(* IEC 61131-3 sources: model-first-plc-agent-ai/results/T3-W-19, 2 files *)

(* ---- a1_code.st ---- *)
FUNCTION_BLOCK TankRuntime
VAR_INPUT
    start : BOOL;
    stop : BOOL;
    LSH : BOOL;
    LSHH : BOOL;
    TON_Duration : TIME;
    TOF_Duration : TIME;
END_VAR
VAR_OUTPUT
    fill_valve : BOOL;
    discharge_valve : BOOL;
END_VAR
VAR
    active_state : INT := 0;
    next_state : INT := 0;
    filling_active : BOOL := FALSE;
    ton_q : BOOL := FALSE;
    tof_q : BOOL := FALSE;
    fill_timer : TON;
    pause_timer : TOF;
END_VAR

(* Evaluate timers using the current GRAFCET situation. *)
filling_active := (active_state = 1);

fill_timer(IN := filling_active, PT := TON_Duration);
pause_timer(IN := filling_active, PT := TOF_Duration);

ton_q := fill_timer.Q;
tof_q := pause_timer.Q;

(* Evaluate transitions from one snapshot of the active situation. *)
next_state := active_state;

CASE active_state OF
    0:
        IF start AND NOT stop AND NOT LSH AND NOT LSHH THEN
            next_state := 1;
        END_IF;

    1:
        IF stop OR LSH OR LSHH THEN
            next_state := 0;
        ELSIF ton_q AND NOT stop AND NOT LSH AND NOT LSHH THEN
            next_state := 2;
        END_IF;

    2:
        IF stop OR LSH OR LSHH THEN
            next_state := 0;
        ELSIF NOT tof_q AND NOT stop AND NOT LSH AND NOT LSHH THEN
            next_state := 1;
        END_IF;

ELSE
    next_state := 0;
END_CASE;

(* Apply the new situation to the timers immediately.
   This resets TON on leaving filling, starts the TOF off-delay
   on that same departure, and asserts TOF on entering filling.
   No further transition is evaluated during this scan. *)
IF next_state <> active_state THEN
    active_state := next_state;
    filling_active := (active_state = 1);

    fill_timer(IN := filling_active, PT := TON_Duration);
    pause_timer(IN := filling_active, PT := TOF_Duration);

    ton_q := fill_timer.Q;
    tof_q := pause_timer.Q;
END_IF;

fill_valve := (active_state = 1);
discharge_valve := FALSE;

END_FUNCTION_BLOCK

PROGRAM Main
VAR
    StartCommand AT %IX100.0 : BOOL;
    StopCommand AT %IX100.1 : BOOL;
    LSH AT %IX100.2 : BOOL;
    LSHH AT %IX100.3 : BOOL;
    FillValve AT %QX100.0 : BOOL;
    DischargeValve AT %QX100.1 : BOOL;
END_VAR
VAR
    (* Configurable commissioning defaults; adjust for the plant. *)
    TON_Duration : TIME := T#5s;
    TOF_Duration : TIME := T#5s;

    start_edge : R_TRIG;
    start : BOOL := FALSE;
    initialized : BOOL := FALSE;
    controller : TankRuntime;
END_VAR

start_edge(CLK := StartCommand);

(* Seed the edge detector without treating a held startup button
   as a new press. *)
IF NOT initialized THEN
    start := FALSE;
    initialized := TRUE;
ELSE
    start := start_edge.Q;
END_IF;

controller(
    start := start,
    stop := StopCommand,
    LSH := LSH,
    LSHH := LSHH,
    TON_Duration := TON_Duration,
    TOF_Duration := TOF_Duration
);

FillValve := controller.fill_valve;
DischargeValve := controller.discharge_valve;

END_PROGRAM

(* ---- a2_code.st ---- *)
FUNCTION_BLOCK FB_TankFilling
VAR_INPUT
    StartCommand : BOOL;
    StopCommand : BOOL;
    LSH : BOOL;
    LSHH : BOOL;
    TON_Duration : TIME;
    TOF_Duration : TIME;
END_VAR
VAR_OUTPUT
    fill_valve : BOOL;
    discharge_valve : BOOL;
END_VAR
VAR
    SequenceState : INT := 0;
    StartEdge : R_TRIG;
    FillingTON : TON;
    FillingTOF : TOF;
    start : BOOL;
    stop : BOOL;
    ton_q : BOOL;
    tof_q : BOOL;
    FillingActive : BOOL;
END_VAR

StartEdge(CLK := StartCommand);
start := StartEdge.Q;
stop := StopCommand;

(* Both standard timers measure filling-step activity. *)
FillingActive := (SequenceState = 1);
FillingTON(IN := FillingActive, PT := TON_Duration);
FillingTOF(IN := FillingActive, PT := TOF_Duration);

ton_q := FillingTON.Q;
tof_q := FillingTOF.Q;

(* Evaluate at most one sequence transition per invocation. *)
IF stop THEN
    SequenceState := 0;
ELSE
    CASE SequenceState OF
        0:
            IF start AND NOT LSH THEN
                SequenceState := 1;
            END_IF;

        1:
            IF LSH THEN
                SequenceState := 0;
            ELSIF ton_q THEN
                SequenceState := 2;
            END_IF;

        2:
            IF LSH THEN
                SequenceState := 0;
            ELSIF NOT tof_q THEN
                SequenceState := 1;
            END_IF;

        ELSE
            SequenceState := 0;
    END_CASE;
END_IF;

fill_valve := (SequenceState = 1);
discharge_valve := FALSE;

(* LSHH is monitored by the plant interface.
   The supplied GRAFCET defines no separate LSHH transition. *)
END_FUNCTION_BLOCK

PROGRAM Main
VAR
    StartCommand AT %IX100.0 : BOOL;
    StopCommand AT %IX100.1 : BOOL;
    LSH AT %IX100.2 : BOOL;
    LSHH AT %IX100.3 : BOOL;
    FillValve AT %QX100.0 : BOOL;
    DischargeValve AT %QX100.1 : BOOL;
END_VAR
VAR
    TankController : FB_TankFilling;
    (* Configurable example presets; set to the required operating values. *)
    TON_Duration : TIME := T#5s;
    TOF_Duration : TIME := T#5s;
END_VAR

TankController(
    StartCommand := StartCommand,
    StopCommand := StopCommand,
    LSH := LSH,
    LSHH := LSHH,
    TON_Duration := TON_Duration,
    TOF_Duration := TOF_Duration
);

FillValve := TankController.fill_valve;
DischargeValve := TankController.discharge_valve;

END_PROGRAM
